// TIA Portal V20 export
Screen "SYSTEM_SETTINGS_2"  1276x673
  ScreenItem "Title_ScreenOverview_X390_Y2" at 390,2 size 510x57  Type=HmiTextBox
  ScreenItem "Line_Header_X0_Y64" at 0,64 size 1276x0  Type=HmiLine
  ScreenItem "Frame_PLC_Diag" at 105,70 size 1070x225  Type=HmiRectangle
  ScreenItem "Title_PLC-Diag" at 107,72 size 442x25  Type=HmiTextBox
  ScreenItem "Text_MAC" at 107,237 size 135x25  Type=HmiTextBox
  ScreenItem "Text_IP" at 467,237 size 135x25  Type=HmiTextBox
  ScreenItem "Text_Subnet" at 467,264 size 135x25  Type=HmiTextBox
  ScreenItem "Text_Point" at 639,237 size 5x25  Type=HmiTextBox
  ScreenItem "Text_Point_1" at 681,237 size 5x25  Type=HmiTextBox
  ScreenItem "Text_Point_2" at 723,237 size 5x25  Type=HmiTextBox
  ScreenItem "Text_Minus" at 268,237 size 5x25  Type=HmiTextBox
  ScreenItem "Text_Minus_1" at 299,237 size 5x25  Type=HmiTextBox
  ScreenItem "Text_Minus_2" at 330,237 size 5x25  Type=HmiTextBox
  ScreenItem "Text_Minus_3" at 361,237 size 5x25  Type=HmiTextBox
  ScreenItem "Text_Minus_4" at 392,237 size 5x25  Type=HmiTextBox
  ScreenItem "Text_MLFB" at 107,129 size 135x25  Type=HmiTextBox
  ScreenItem "Text_Firmware" at 107,210 size 135x25  Type=HmiTextBox
  ScreenItem "Text_Hardware" at 107,183 size 135x25  Type=HmiTextBox
  ScreenItem "Text_SerialNo" at 107,156 size 135x25  Type=HmiTextBox
  ScreenItem "Text_InstallationDate" at 827,209 size 135x25  Type=HmiTextBox
  ScreenItem "Text_AddInfo" at 827,236 size 135x25  Type=HmiTextBox
  ScreenItem "Text_PlantDesignation" at 827,102 size 160x25  Type=HmiTextBox
  ScreenItem "Text_ManufacturerID" at 107,102 size 135x25  Type=HmiTextBox
  ScreenItem "Text_RevisionCount" at 467,102 size 135x25  Type=HmiTextBox
  ScreenItem "Text_ProfileID" at 467,129 size 135x25  Type=HmiTextBox
  ScreenItem "Text_ProfileSpec" at 467,156 size 135x25  Type=HmiTextBox
  ScreenItem "Text_IMVersion" at 467,183 size 135x25  Type=HmiTextBox
  ScreenItem "Text_IMSupported" at 467,210 size 135x25  Type=HmiTextBox
  ScreenItem "ManufacturerID" at 243,102 size 65x25  Type=HmiIOField
  ScreenItem "MLFB" at 243,129 size 220x25  Type=HmiIOField
  ScreenItem "MLFB_1" at 243,156 size 220x25  Type=HmiIOField
  ScreenItem "Hardware" at 243,183 size 65x25  Type=HmiIOField
  ScreenItem "FirmwareType" at 243,210 size 24x25  Type=HmiIOField
  ScreenItem "FirmwareFunctional" at 274,210 size 24x25  Type=HmiIOField
  ScreenItem "Text_Point_3" at 299,210 size 5x25  Type=HmiTextBox
  ScreenItem "FirmwareBugfix" at 305,210 size 24x25  Type=HmiIOField
  ScreenItem "Text_Point_7" at 330,210 size 5x25  Type=HmiTextBox
  ScreenItem "FirmwareInternal" at 336,210 size 24x25  Type=HmiIOField
  ScreenItem "Mac1" at 243,237 size 24x25  Type=HmiIOField
  ScreenItem "Mac2" at 274,237 size 24x25  Type=HmiIOField
  ScreenItem "Mac3" at 305,237 size 24x25  Type=HmiIOField
  ScreenItem "Mac4" at 336,237 size 24x25  Type=HmiIOField
  ScreenItem "Mac5" at 367,237 size 24x25  Type=HmiIOField
  ScreenItem "Mac6" at 398,237 size 24x25  Type=HmiIOField
  ScreenItem "RevisionCount" at 603,102 size 60x25  Type=HmiIOField
  ScreenItem "ProfileID" at 603,129 size 60x25  Type=HmiIOField
  ScreenItem "ProfileSpec" at 603,156 size 60x25  Type=HmiIOField
  ScreenItem "IMVersion" at 603,183 size 60x25  Type=HmiIOField
  ScreenItem "IMSupported" at 603,210 size 60x25  Type=HmiIOField
  ScreenItem "IP1" at 603,237 size 35x25  Type=HmiIOField
  ScreenItem "IP2" at 645,237 size 35x25  Type=HmiIOField
  ScreenItem "IP3" at 687,237 size 35x25  Type=HmiIOField
  ScreenItem "IP4" at 729,237 size 35x25  Type=HmiIOField
  ScreenItem "PlantDesignation" at 827,129 size 342x25  Type=HmiIOField
  ScreenItem "InstallationDate" at 963,209 size 206x25  Type=HmiIOField
  ScreenItem "AddInfo" at 827,262 size 342x27  Type=HmiIOField
  ScreenItem "Text_Point_4" at 639,264 size 5x25  Type=HmiTextBox
  ScreenItem "Text_Point_5" at 681,264 size 5x25  Type=HmiTextBox
  ScreenItem "Text_Point_6" at 723,264 size 5x25  Type=HmiTextBox
  ScreenItem "Subnet1" at 603,264 size 35x25  Type=HmiIOField
  ScreenItem "Subnet2" at 645,264 size 35x25  Type=HmiIOField
  ScreenItem "Subnet3" at 687,264 size 35x25  Type=HmiIOField
  ScreenItem "Subnet4" at 729,264 size 35x25  Type=HmiIOField
  ScreenItem "Text_LocationIdentifier" at 827,154 size 160x25  Type=HmiTextBox
  ScreenItem "LocationIdentifier" at 827,181 size 342x25  Type=HmiIOField
  ScreenItem "Button_UpdateIuM" at 1,70 size 90x60  Type=HmiButton
  ScreenItem "Button_SystemSettings" at 95,2 size 90x60  Type=HmiButton
  ScreenItem "Button_SICARHelp" at 1183,2 size 90x60  Type=HmiButton
  ScreenItem "permanentareaborderrectangle" at 0,0 size 0x0  Type=HmiRectangle
  ScreenItem "Button_Back" at 2,2 size 90x60  Type=HmiButton
